// TwinCAT 3 PLC project PLC_ValveCharact
// ProgramVersion: 3.1.4026.30
// libraries:
//   Tc2_Standard, * (Beckhoff Automation GmbH)
//   Tc2_System, * (Beckhoff Automation GmbH)
//   Tc3_Mc3FluidPower, * (Beckhoff Automation GmbH)
//   Tc3_Mc3Ptp, * (Beckhoff Automation GmbH)
// project tree:
//   / MC_Task_MET_.TcTTO, PlcTask.TcTTO
//   POUs/ MAIN.TcPOU, Simu.TcPOU
// real-time tasks:
//   TASK Job Task: cycle default, priority 32
//   TASK MC-Task (MET): cycle T#2ms, priority 3, ADS port 521
//   TASK MC-Task (MPT): cycle T#10ms, priority 8, ADS port 531
//   TASK PlcTask: cycle T#10ms, priority 20, ADS port 350
// variable links:
//   PLC_ValveCharact/PLC_ValveCharact Instance <-> MC Project1/Axes/Axis
//     MC_Task_MET_ Inputs/Simu.SetVelo <-> Analog Outputs/Output
//     MC_Task_MET_ Outputs/Simu.ActPos <-> SSI Inputs/Counter Value
//     PlcTask Inputs/MAIN.HydAxis.McToPlc/Act <-> McToPlc/Act
//     PlcTask Inputs/MAIN.HydAxis.McToPlc/Set <-> McToPlc/Set
//     PlcTask Inputs/MAIN.HydAxis.McToPlc/Std <-> McToPlc/Std
//     PlcTask Outputs/MAIN.HydAxis.PlcToMc/Std <-> PlcToMc/Std
//   PLC_ValveCharact/PLC_ValveCharact Instance <-> MC Project1/Axes/Axis/Pressure Sensor A
//     PlcTask Outputs/Simu.PressureA <-> Analog Inputs/Counter Value
//   PLC_ValveCharact/PLC_ValveCharact Instance <-> MC Project1/Axes/Axis/Valve Characteristic Curve
//     PlcTask Inputs/MAIN.fbValveObject.McToPlc/Oid <-> McToPlc/Oid

CONFIGURATION PLC_ValveCharact
    RESOURCE PLC ON TwinCAT3
        TASK MC_Task_MET_(INTERVAL := T#2ms, PRIORITY := 3);
        TASK PlcTask(INTERVAL := T#10ms, PRIORITY := 20);
        PROGRAM Simu WITH MC_Task_MET_ : Simu;
        PROGRAM MAIN WITH PlcTask : MAIN;
    END_RESOURCE
END_CONFIGURATION

// ---- POUs/Simu.TcPOU
// Simulation program for the Valve Characterization sample.
// Models a non-linear hydraulic valve: integrates the (non-linear) spool velocity to an actual
// position and feeds simulated I/O, so the sample runs without real hardware.
PROGRAM Simu
VAR
	ActPos AT%Q*:	DINT;
	SetVelo AT%I*:	INT;
	PressureA AT%Q*:	INT;
 
 	fSetVelo:	LREAL;
 	fActPos:	LREAL;

	fSetVeloNonLinear: LREAL;
END_VAR


fSetVelo:=INT_TO_LREAL(SetVelo)/32767*500.0;

IF fSetVelo > 0.0 THEN
	fSetVeloNonLinear := (1-COS(fSetVelo/500.0*3.14))/2.0*500.0;
ELSE
	fSetVeloNonLinear := -(1-COS(fSetVelo/500.0*3.14))/2.0*500.0;
END_IF
//fSetVeloNonLinear:=fSetVelo;
fActPos:=fActPos+fSetVeloNonLinear*0.002;

fActPos:=MIN(MAX(fActPos,0.0),500.0);
ActPos:=LREAL_TO_DINT(fActPos * 1000.0);

END_PROGRAM

// ---- POUs/MAIN.TcPOU
// Valve Characterization sample
// Shows automated valve characterization (spool position -> axis velocity) using
// MC_ValveCharacterization and MC_ValveCharacteristicCurve; the separate Simu program models a
// non-linear valve so the sample runs without hardware.
// Operation: set bStart := TRUE to power, traverse and characterize; then use bEnable/bDisable/bReadValveCharacteristicCurve.
PROGRAM MAIN
VAR
	bStart: 							BOOL;
	bEnableValveCharacteristicCurve: 	BOOL;
	bDisableValveCharacteristicCurve: 	BOOL;
	bReadValveCharacteristicCurve:		BOOL;
	nNumberOfValveCharacteristicCurvePoints:	UDINT:=21;

	nErrorId:		UDINT;

	HydAxis:			AXIS_REF;
	fbPower:			MC_Power;
	
	fbValveObject:			MC_ValveCharacteristicCurve;
	fbCharacterization:		MC_ValveCharacterization;
	stValveCharactOptions:	ValveCharacterizationOptions;
	
	fbMoveAbsFwd:		MC_MoveAbsolute;
	fbMoveAbsBwd:		MC_MoveAbsolute;
	fbTimer:				TON;	
	
	nNoOfPoints:		UDINT;
	i:				INT;
	aValvePoint:		ARRAY[1..cnNumberOfValveCharacteristicCurvePoints] OF ValveCharacteristicPoint;
	
	bInit: 			BOOL;
	nState: 		INT;
	
	fXValue:		LREAL;
	fYValue:		LREAL;
END_VAR
VAR CONSTANT
	cnNumberOfValveCharacteristicCurvePoints:		UDINT:=100;
END_VAR

nNumberOfValveCharacteristicCurvePoints := MIN(cnNumberOfValveCharacteristicCurvePoints, nNumberOfValveCharacteristicCurvePoints);

IF bStart THEN
	fbPower.Enable:=TRUE;
END_IF
fbPower
(
	Axis:=HydAxis,
	EnableNegative:=TRUE,
	EnablePositive:=TRUE
);

IF NOT bInit AND fbPower.Status AND 0 = nErrorId THEN
	nErrorId := fbValveObject.Connect();
	bInit:= fbValveObject.IsConnected;
END_IF


CASE nState OF
	0:
	IF bStart AND fbValveObject.IsConnected THEN
		fbValveObject.Disable();
		nState:=nState+1;
	END_IF
	

	1:
	IF fbPower.Status THEN
		fbMoveAbsFwd.Position:=250.0;
		fbMoveAbsFwd.Velocity:=500.0;
		fbMoveAbsFwd.Execute:=TRUE;
		bStart:=FALSE;
		nState:=nState+1;
	END_IF

	2:
	IF NOT fbMoveAbsFwd.Busy THEN
		fbMoveAbsFwd.Execute:=FALSE;		
		IF fbMoveAbsFwd.Done THEN	
			fbMoveAbsBwd.Position:=0.0;
			fbMoveAbsBwd.Velocity:=500.0;
			fbMoveAbsBwd.Execute:=TRUE;		
			nState:=nState+1;
		END_IF
	END_IF
	
	3:
	IF NOT fbMoveAbsBwd.Busy THEN
		fbMoveAbsBwd.Execute:=FALSE;		
		IF fbMoveAbsBwd.Done THEN	
			fbTimer.PT:=T#1S;
			fbTimer.IN:=TRUE;
			nState:=nState+1;
		END_IF
	END_IF
	
	4:
	IF fbTimer.Q THEN
		fbTimer.IN:=FALSE;
		fbCharacterization.Execute:=TRUE;
		nState:=nState+1;
	END_IF


	5:
	IF NOT fbCharacterization.Busy THEN
		IF fbCharacterization.Done THEN
			fbCharacterization.Execute:=FALSE;
			fbValveObject.Enable();
			fbTimer.IN:=TRUE;
			nState:=nState+1;
		END_IF
	END_IF

	6:
		nState:=nState+1;

	7:
	IF fbTimer.Q THEN			
		fbMoveAbsFwd.Position:=250.0;
		fbMoveAbsFwd.Velocity:=500.0;
		fbMoveAbsFwd.Execute:=TRUE;
		fbTimer.IN:=FALSE;
			nState:=nState+1;
	END_IF

	8:
	IF NOT fbMoveAbsFwd.Busy THEN
		fbMoveAbsFwd.Execute:=FALSE;		
		IF fbMoveAbsFwd.Done THEN	
			fbMoveAbsBwd.Position:=0.0;
			fbMoveAbsBwd.Velocity:=500.0;
			fbMoveAbsBwd.Execute:=TRUE;		
			nState:=nState+1;
		END_IF
	END_IF
	
	9:
	IF NOT fbMoveAbsBwd.Busy THEN
		fbMoveAbsBwd.Execute:=false;		
		IF fbMoveAbsBwd.Done THEN	
			nState:=0;
		END_IF
	END_IF
END_CASE

fbTimer();

stValveCharactOptions.MinimumTravelPerMeasurement:=0.2;
stValveCharactOptions.WaitTimeAfterVelocityStep:=0.1;
stValveCharactOptions.WaitTimeAtPositionLimit:=0.2;
stValveCharactOptions.OutputLimit:=1.0;
fbCharacterization
(
	Axis:=HydAxis,
	OutputStepsize:=2.0/TO_LREAL(nNumberOfValveCharacteristicCurvePoints - 1),
	PositionLimitMinimum:=50.0,
	PositionLimitMaximum:=450.0,
	Options:=stValveCharactOptions
);


IF bReadValveCharacteristicCurve THEN
	nNoOfPoints:=nNumberOfValveCharacteristicCurvePoints;
	fbValveObject.ReadData(DestinationAddress:=ADR(aValvePoint), NumberOfPoints:=nNoOfPoints);
	
	i:=i+1;
	IF i > nNoOfPoints THEN
		i:=1;
	END_IF
	fXValue := aValvePoint[i].SpoolPosition;
	fYValue := aValvePoint[i].Velocity;
END_IF




IF bEnableValveCharacteristicCurve THEN
	nErrorId := fbValveObject.Enable();
	bEnableValveCharacteristicCurve:=FALSE;
END_IF

IF bDisableValveCharacteristicCurve THEN
	nErrorId := fbValveObject.Disable();
	bDisableValveCharacteristicCurve:=FALSE;
END_IF


fbMoveAbsFwd
(
	Axis:=HydAxis,
);

fbMoveAbsBwd
(
	Axis:=HydAxis,
);

END_PROGRAM
